Fanuc KAREL source: KA00112.KL

PROGRAM KA00112
%NOLOCKGROUP
VAR
  SRC: CONFIG
  DST: STRING[80]
BEGIN
  SRC.CFG_FLIP = TRUE
  DST = SRC
END KA00112
